ADAPTER mgz_sensor (* Adapter Interface *)
  (* Standard: 61499-1 *)
  (* Version 0.0, 10/27/2026, lizar, Schneider Electric *)
  PACKAGE Main;
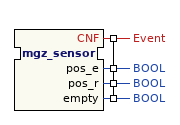
  EVENT_OUTPUT
    CNF WITH pos_e, pos_r, empty; (* Confirmation from Plug *)
  END_EVENT
  VAR_OUTPUT
    pos_e : BOOL;
    pos_r : BOOL;
    empty : BOOL;
  END_VAR
  SERVICE SOCKET/PLUG
    SEQUENCE request_confirm
      SOCKET.REQ(REQD) -> PLUG.REQ(REQD);
      PLUG.CNF(CNFD) -> SOCKET.CNF(CNFD);
    END_SEQUENCE
    SEQUENCE indication_response
      PLUG.IND(INDD) -> SOCKET.IND(INDD);
      SOCKET.RSP(RSPD) -> PLUG.RSP(RSPD);
    END_SEQUENCE
  END_SERVICE
END_ADAPTER
